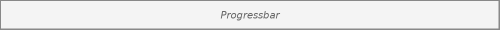
VISUALIZATION vis_ProgressBar  // 500x30
    Progressbar (0,0 500x30), variable: g_HMI_Panel.stPLC_To_VisuPLC.fBlendingPercenatge
END_VISUALIZATION

(* stored: Version 1.1.0.1, ProductVersion 3.1.4024.15
   Visu vis_ProgressBar: Id {4d1ad0d8-54bb-4713-aa1d-c39318435f7f} *)
